FUNCTION "LGF_BinaryMaskCompare" : Bool
{ S7_Optimized_Access := 'TRUE' }
AUTHOR : Siemens_Simatic_Systems_Support
FAMILY : LGF
NAME : LGF_BinaryMaskCompare
   VAR_INPUT
      source : DWord;
      compare : DWord;
      mask { S7_PredefinedAssignment := '16#FFFFFFFF'; S7_HiddenAssignment := 'Show'; S7_ShowAssignmentIfParamsNotIdentical := 'false'} : DWord;
   END_VAR

   VAR CONSTANT
      ALL_BITS_ARE_FALSE : DWord := 16#00000000;
   END_VAR


BEGIN
	REGION BLOCK INFO HEADER
	  //===============================================================================
	  // SIEMENS AG / (c)Copyright 2019
	  //-------------------------------------------------------------------------------
	  // Title:            LGF_BinaryMaskCompare
	  // Comment/Function: Comparing two binary Values `source` and `compare` by a given `mask`.
	  //                   Both given values are masked, and the results is than compared and returned
	  //                   Can be used for Word and Byte as well, by convert the passed parameter using for e.g. Byte_to_DWord(...)
	  // Library/Family:   LGF (Library General Functions)
	  // Author:           Siemens Simatic Systems Support
	  // Tested with:      1516F FW2.8 / S7-PLCSIM Advanced V3.0
	  // Engineering:      TIA Portal V16 Update 4
	  // Restrictions:     ENO not in use, set to true, no error handling
	  // Requirements:     PLC (S7-1200 / S7-1500)
	  //-------------------------------------------------------------------------------
	  //===============================================================================
	END_REGION BLOCK INFO HEADER

	//Mask Compare Equal DWord
	#LGF_BinaryMaskCompare := (((#source AND #mask) XOR (#compare AND #mask)) = #ALL_BITS_ARE_FALSE);

	// ENO is not used, forced to TRUE
	ENO := TRUE;

END_FUNCTION